// SIMATIC S7-200 project (STEP 7-Micro/WIN), CPU 226 CN REL 02.01

SYMBOL_TABLE 用户定义1
原点传感器检测          I0.0
右限位行程开关          I0.1
左限位行程开关          I0.2
机械手抬升下限检测        I0.3
机械手抬升上限检测        I0.4
机械手旋转左旋检测        I0.5
机械手旋转右旋检测        I0.6
机械手伸出检测          I0.7
机械手缩回检测          I1.0
机械手夹紧检测          I1.1
伺服报警             I1.2
按钮SB2            I2.4
按钮SB1            I2.5
急停               I2.6
全线速度             I2.7
初始状态检查           M0.0
回原点开始            M0.1
回原点完成            M0.2
正向点动             M0.3
反向点动             M0.4
双按键              M0.5
网络正常             M1.0
全线模式             M1.1
机械手复位            M1.2
准备就绪             M1.3
全线启动             M1.4
全线停止             M1.5
脉冲               Q0.0
方向               Q0.1
提升台上升电磁阀         Q0.3
回转气缸左旋电磁阀        Q0.4
回转气缸右旋电磁阀        Q0.5
手爪伸出电磁阀          Q0.6
手爪夹紧电磁阀          Q0.7
手爪放松电磁阀          Q1.0
黄色指示灯            Q1.5
绿色指示灯            Q1.6
红色指示灯            Q1.7
测试开始             S1.0
复位               V100.0
启动               V100.1
初始状态指示           V200.0
确认保存             V200.1
测试完成             V200.2
运行模式             V200.5
允许返回             V200.6
自动返回             V200.7
绿色警示灯            V1000.0
黄色警示灯            V1000.1
红色警示灯            V1000.2
各站红灯             V1000.3
供料请求             V1000.4
允许装配             V1000.5
允许加工             V1000.6
允许分拣             V1000.7
料不足_供料           V1020.2
缺料_供料            V1020.3
供料完成             V1020.4
料不足_装配           V1030.2
缺料_装配            V1030.3
装配完成             V1030.4
装配急停             V1030.5
故障无法修复           V1030.6
加工完成             V1040.2
停止完成             V1050.2
测试项              VB110
计划生产套件数          VB120
已生产套件数           VB1051
供料站位置            VD210
装配站位置            VD220
加工站位置            VD230
分拣站位置            VD240
当前绝对位置           VD250
当前速度             VD260
停止               V1001.0
END_SYMBOL_TABLE

ORGANIZATION_BLOCK 主程序:OB1
TITLE=程序注释
BEGIN
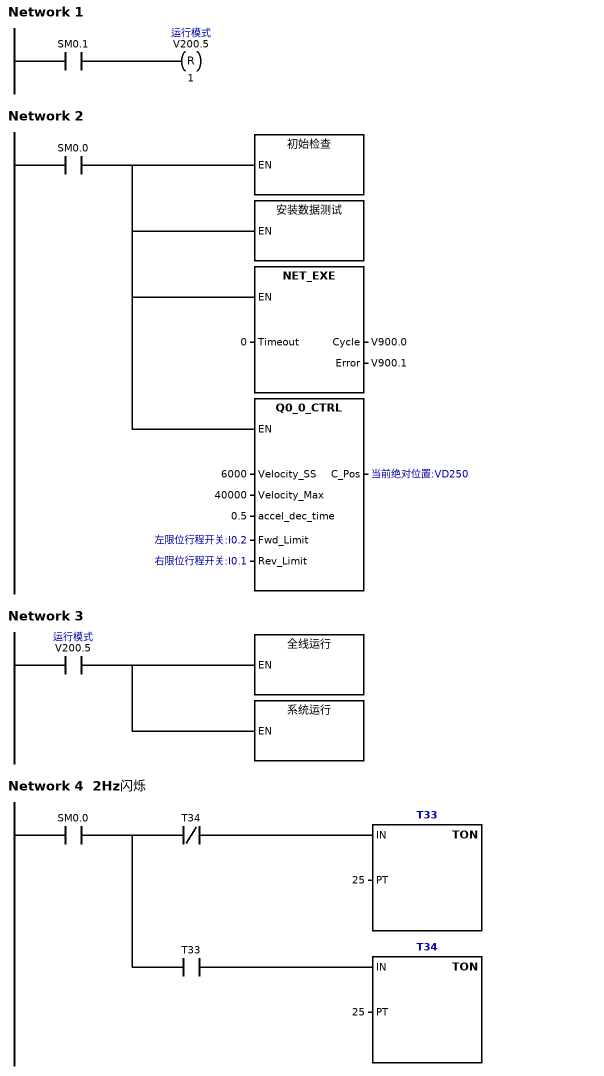
Network 1
LD     SM0.1
R      运行模式:V200.5, 1
Network 2
LD     SM0.0
CALL   初始检查:SBR0
CALL   安装数据测试:SBR8
CALL   NET_EXE:SBR11, 0, V900.0, V900.1
CALL   Q0_0_CTRL:SBR1, 6000, 40000, 0.5, 左限位行程开关:I0.2, 右限位行程开关:I0.1, 当前绝对位置:VD250
Network 3
LD     运行模式:V200.5
CALL   全线运行:SBR13
CALL   系统运行:SBR14
Network 4 // 2Hz闪烁
LD     SM0.0
LPS
AN     T34
TON    T33, 25
LPP
A      T33
TON    T34, 25
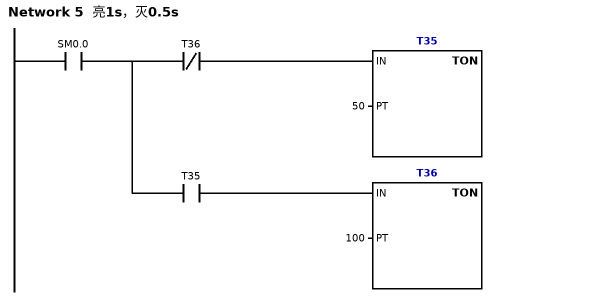
Network 5 // 亮1s，灭0.5s
LD     SM0.0
LPS
AN     T36
TON    T35, 50
LPP
A      T35
TON    T36, 100
END_ORGANIZATION_BLOCK

SUBROUTINE_BLOCK 初始检查:SBR0
TITLE=子程序注释
BEGIN
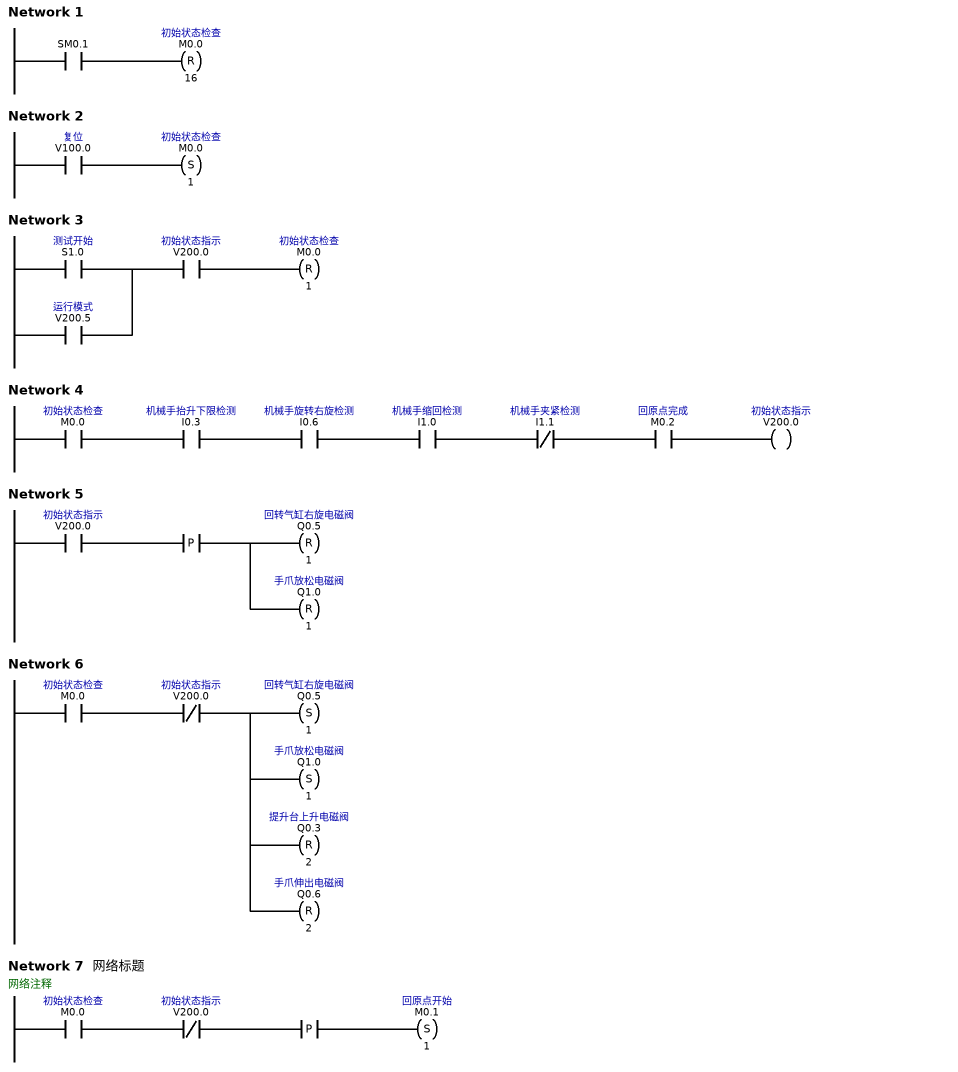
Network 1
LD     SM0.1
R      初始状态检查:M0.0, 16
Network 2
LD     复位:V100.0
S      初始状态检查:M0.0, 1
Network 3
LD     测试开始:S1.0
O      运行模式:V200.5
A      初始状态指示:V200.0
R      初始状态检查:M0.0, 1
Network 4
LD     初始状态检查:M0.0
A      机械手抬升下限检测:I0.3
A      机械手旋转右旋检测:I0.6
A      机械手缩回检测:I1.0
AN     机械手夹紧检测:I1.1
A      回原点完成:M0.2
=      初始状态指示:V200.0
Network 5
LD     初始状态指示:V200.0
EU
R      回转气缸右旋电磁阀:Q0.5, 1
R      手爪放松电磁阀:Q1.0, 1
Network 6
LD     初始状态检查:M0.0
AN     初始状态指示:V200.0
S      回转气缸右旋电磁阀:Q0.5, 1
S      手爪放松电磁阀:Q1.0, 1
R      提升台上升电磁阀:Q0.3, 2
R      手爪伸出电磁阀:Q0.6, 2
Network 7 // 网络标题
// 网络注释
LD     初始状态检查:M0.0
AN     初始状态指示:V200.0
EU
S      回原点开始:M0.1, 1
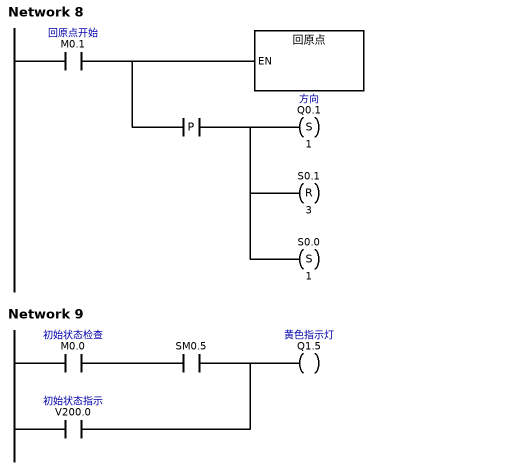
Network 8
LD     回原点开始:M0.1
CALL   回原点:SBR7
EU
S      方向:Q0.1, 1
R      S0.1, 3
S      S0.0, 1
Network 9
LD     初始状态检查:M0.0
A      SM0.5
O      初始状态指示:V200.0
=      黄色指示灯:Q1.5
END_SUBROUTINE_BLOCK

// SBR1: protected block, not included

// SBR2: protected block, not included

// SBR3: protected block, not included

// SBR4: protected block, not included

// SBR5: protected block, not included

// SBR6: protected block, not included

SUBROUTINE_BLOCK 回原点:SBR7
TITLE=子程序注释
BEGIN
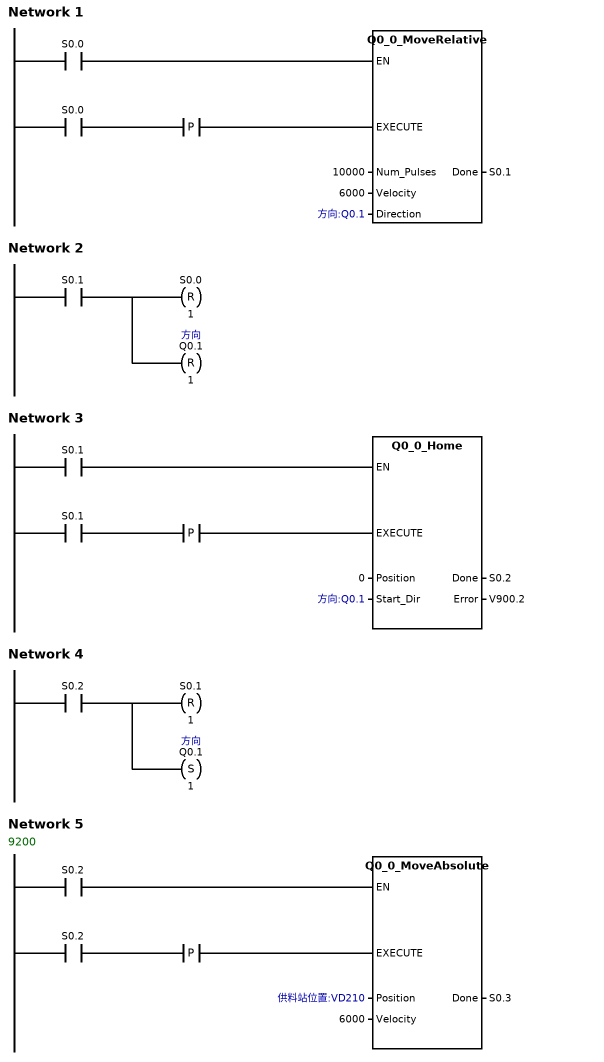
Network 1
LD     S0.0
=      L60.0
LD     S0.0
EU
=      L63.7
LD     L60.0
CALL   Q0_0_MoveRelative:SBR3, L63.7, 10000, 6000, 方向:Q0.1, S0.1
Network 2
LD     S0.1
R      S0.0, 1
R      方向:Q0.1, 1
Network 3
LD     S0.1
=      L60.0
LD     S0.1
EU
=      L63.7
LD     L60.0
CALL   Q0_0_Home:SBR5, L63.7, 0, 方向:Q0.1, S0.2, V900.2
Network 4
LD     S0.2
R      S0.1, 1
S      方向:Q0.1, 1
Network 5
// 9200
LD     S0.2
=      L60.0
LD     S0.2
EU
=      L63.7
LD     L60.0
CALL   Q0_0_MoveAbsolute:SBR4, L63.7, 供料站位置:VD210, 6000, S0.3
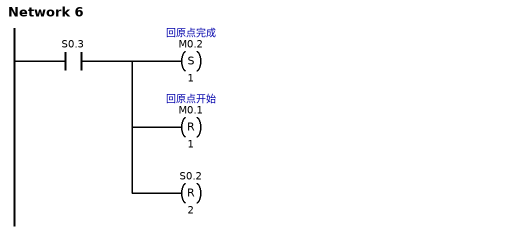
Network 6
LD     S0.3
S      回原点完成:M0.2, 1
R      回原点开始:M0.1, 1
R      S0.2, 2
Network 7 // 网络标题
// 网络注释
Network 9 // 网络标题
// 网络注释
END_SUBROUTINE_BLOCK

SUBROUTINE_BLOCK 安装数据测试:SBR8
TITLE=子程序注释
BEGIN
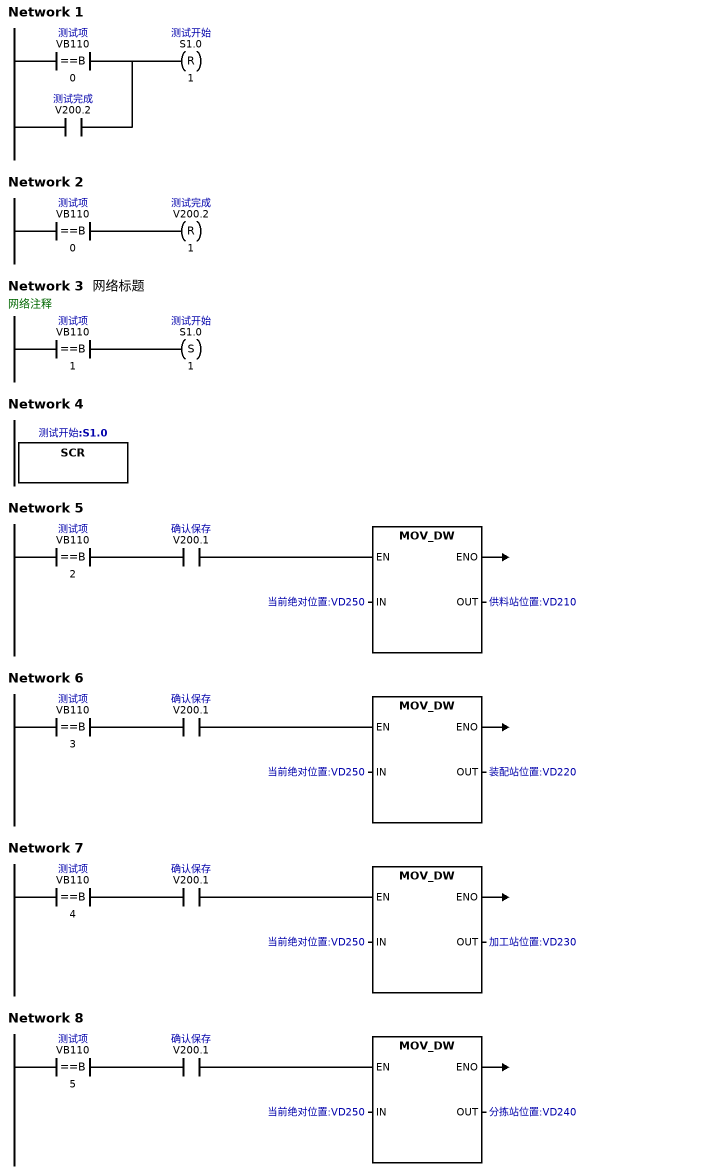
Network 1
LDB=   测试项:VB110, 0
O      测试完成:V200.2
R      测试开始:S1.0, 1
Network 2
LDB=   测试项:VB110, 0
R      测试完成:V200.2, 1
Network 3 // 网络标题
// 网络注释
LDB=   测试项:VB110, 1
S      测试开始:S1.0, 1
Network 4
LSCR   测试开始:S1.0
Network 5
LDB=   测试项:VB110, 2
A      确认保存:V200.1
MOVD   当前绝对位置:VD250, 供料站位置:VD210
Network 6
LDB=   测试项:VB110, 3
A      确认保存:V200.1
MOVD   当前绝对位置:VD250, 装配站位置:VD220
Network 7
LDB=   测试项:VB110, 4
A      确认保存:V200.1
MOVD   当前绝对位置:VD250, 加工站位置:VD230
Network 8
LDB=   测试项:VB110, 5
A      确认保存:V200.1
MOVD   当前绝对位置:VD250, 分拣站位置:VD240
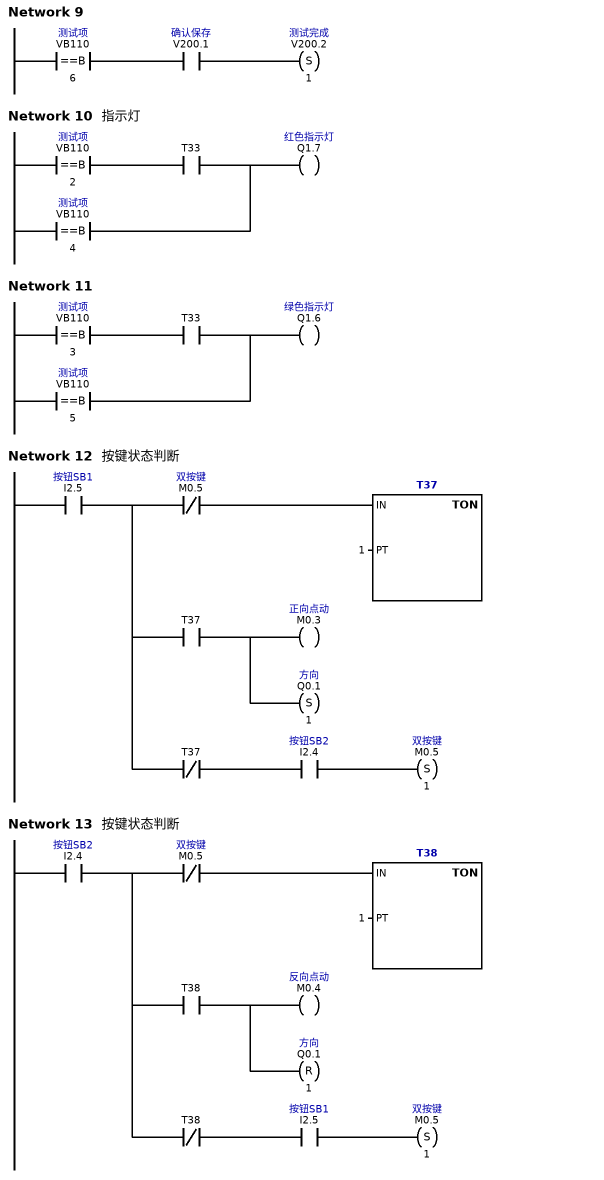
Network 9
LDB=   测试项:VB110, 6
A      确认保存:V200.1
S      测试完成:V200.2, 1
Network 10 // 指示灯
LDB=   测试项:VB110, 2
A      T33
OB=    测试项:VB110, 4
=      红色指示灯:Q1.7
Network 11
LDB=   测试项:VB110, 3
A      T33
OB=    测试项:VB110, 5
=      绿色指示灯:Q1.6
Network 12 // 按键状态判断
LD     按钮SB1:I2.5
LPS
AN     双按键:M0.5
TON    T37, 1
LRD
A      T37
=      正向点动:M0.3
S      方向:Q0.1, 1
LPP
AN     T37
A      按钮SB2:I2.4
S      双按键:M0.5, 1
Network 13 // 按键状态判断
LD     按钮SB2:I2.4
LPS
AN     双按键:M0.5
TON    T38, 1
LRD
A      T38
=      反向点动:M0.4
R      方向:Q0.1, 1
LPP
AN     T38
A      按钮SB1:I2.5
S      双按键:M0.5, 1
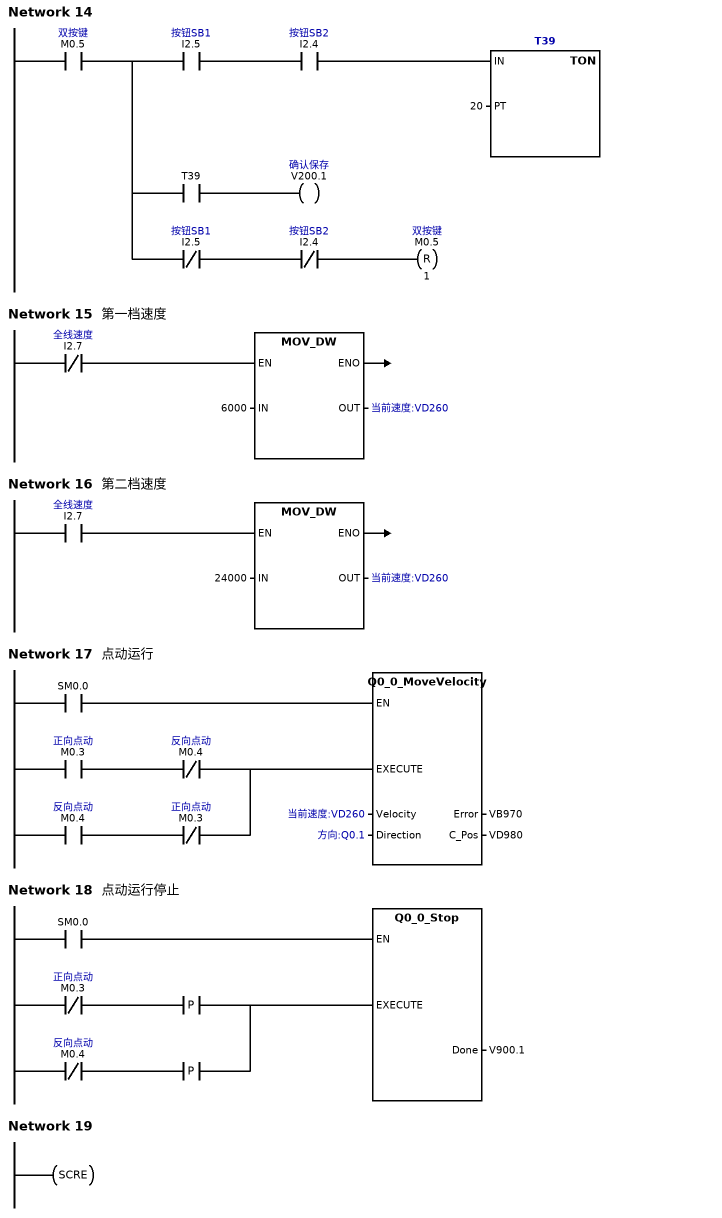
Network 14
LD     双按键:M0.5
LPS
A      按钮SB1:I2.5
A      按钮SB2:I2.4
TON    T39, 20
LRD
A      T39
=      确认保存:V200.1
LPP
AN     按钮SB1:I2.5
AN     按钮SB2:I2.4
R      双按键:M0.5, 1
Network 15 // 第一档速度
LDN    全线速度:I2.7
MOVD   6000, 当前速度:VD260
Network 16 // 第二档速度
LD     全线速度:I2.7
MOVD   24000, 当前速度:VD260
Network 17 // 点动运行
LD     SM0.0
=      L60.0
LD     正向点动:M0.3
AN     反向点动:M0.4
LD     反向点动:M0.4
AN     正向点动:M0.3
OLD
=      L63.7
LD     L60.0
CALL   Q0_0_MoveVelocity:SBR9, L63.7, 当前速度:VD260, 方向:Q0.1, VB970, VD980
Network 18 // 点动运行停止
LD     SM0.0
=      L60.0
LDN    正向点动:M0.3
EU
LDN    反向点动:M0.4
EU
OLD
=      L63.7
LD     L60.0
CALL   Q0_0_Stop:SBR10, L63.7, V900.1
Network 19
SCRE
END_SUBROUTINE_BLOCK

// SBR9: protected block, not included

// SBR10: protected block, not included

// SBR11: protected block, not included

SUBROUTINE_BLOCK 全线运行:SBR13
TITLE=
BEGIN
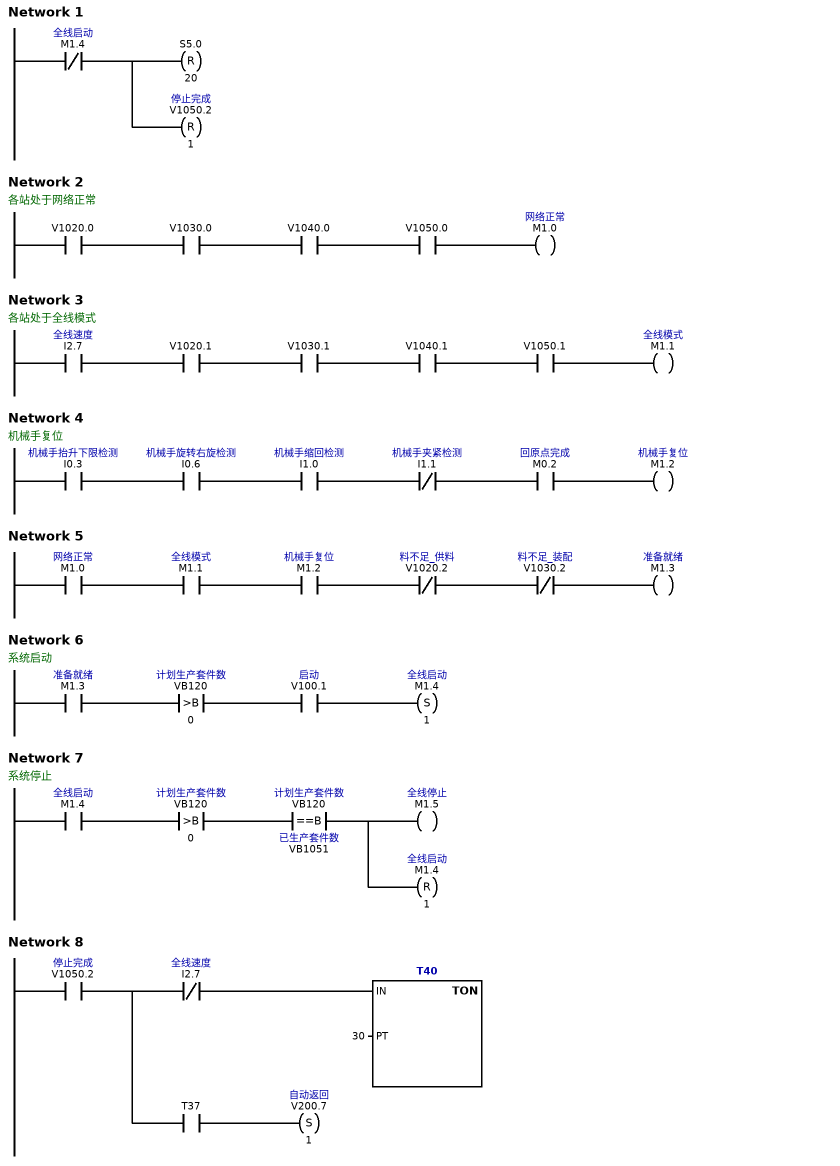
Network 1
LDN    全线启动:M1.4
R      S5.0, 20
R      停止完成:V1050.2, 1
Network 2
// 各站处于网络正常
LD     V1020.0
A      V1030.0
A      V1040.0
A      V1050.0
=      网络正常:M1.0
Network 3
// 各站处于全线模式
LD     全线速度:I2.7
A      V1020.1
A      V1030.1
A      V1040.1
A      V1050.1
=      全线模式:M1.1
Network 4
// 机械手复位
LD     机械手抬升下限检测:I0.3
A      机械手旋转右旋检测:I0.6
A      机械手缩回检测:I1.0
AN     机械手夹紧检测:I1.1
A      回原点完成:M0.2
=      机械手复位:M1.2
Network 5
LD     网络正常:M1.0
A      全线模式:M1.1
A      机械手复位:M1.2
AN     料不足_供料:V1020.2
AN     料不足_装配:V1030.2
=      准备就绪:M1.3
Network 6
// 系统启动
LD     准备就绪:M1.3
AB>    计划生产套件数:VB120, 0
A      启动:V100.1
S      全线启动:M1.4, 1
Network 7
// 系统停止
LD     全线启动:M1.4
AB>    计划生产套件数:VB120, 0
AB=    计划生产套件数:VB120, 已生产套件数:VB1051
=      全线停止:M1.5
R      全线启动:M1.4, 1
Network 8
LD     停止完成:V1050.2
LPS
AN     全线速度:I2.7
TON    T40, 30
LPP
A      T37
S      自动返回:V200.7, 1
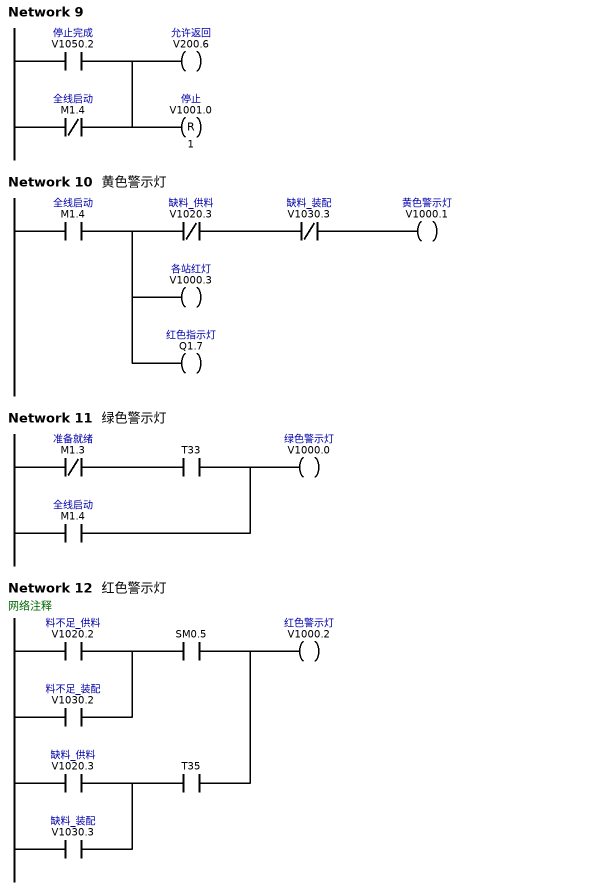
Network 9
LD     停止完成:V1050.2
ON     全线启动:M1.4
=      允许返回:V200.6
R      停止:V1001.0, 1
Network 10 // 黄色警示灯
LD     全线启动:M1.4
LPS
AN     缺料_供料:V1020.3
AN     缺料_装配:V1030.3
=      黄色警示灯:V1000.1
LRD
=      各站红灯:V1000.3
LPP
=      红色指示灯:Q1.7
Network 11 // 绿色警示灯
LDN    准备就绪:M1.3
A      T33
O      全线启动:M1.4
=      绿色警示灯:V1000.0
Network 12 // 红色警示灯
// 网络注释
LD     料不足_供料:V1020.2
O      料不足_装配:V1030.2
A      SM0.5
LD     缺料_供料:V1020.3
O      缺料_装配:V1030.3
A      T35
OLD
=      红色警示灯:V1000.2
END_SUBROUTINE_BLOCK

SUBROUTINE_BLOCK 系统运行:SBR14
TITLE=子程序注释
BEGIN
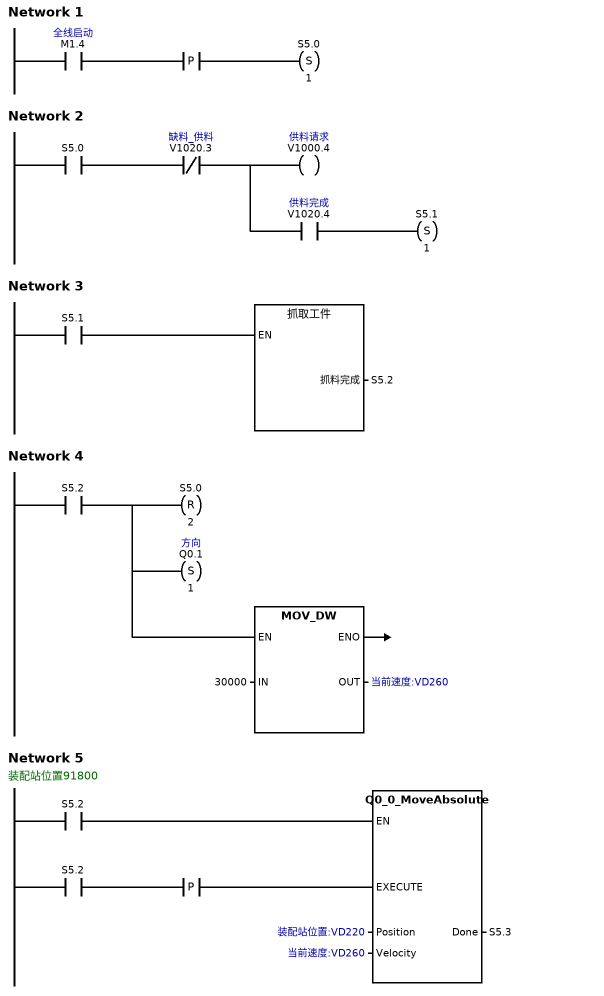
Network 1
LD     全线启动:M1.4
EU
S      S5.0, 1
Network 2
LD     S5.0
AN     缺料_供料:V1020.3
=      供料请求:V1000.4
A      供料完成:V1020.4
S      S5.1, 1
Network 3
LD     S5.1
CALL   抓取工件:SBR15, S5.2
Network 4
LD     S5.2
R      S5.0, 2
S      方向:Q0.1, 1
MOVD   30000, 当前速度:VD260
Network 5
// 装配站位置91800
LD     S5.2
=      L60.0
LD     S5.2
EU
=      L63.7
LD     L60.0
CALL   Q0_0_MoveAbsolute:SBR4, L63.7, 装配站位置:VD220, 当前速度:VD260, S5.3
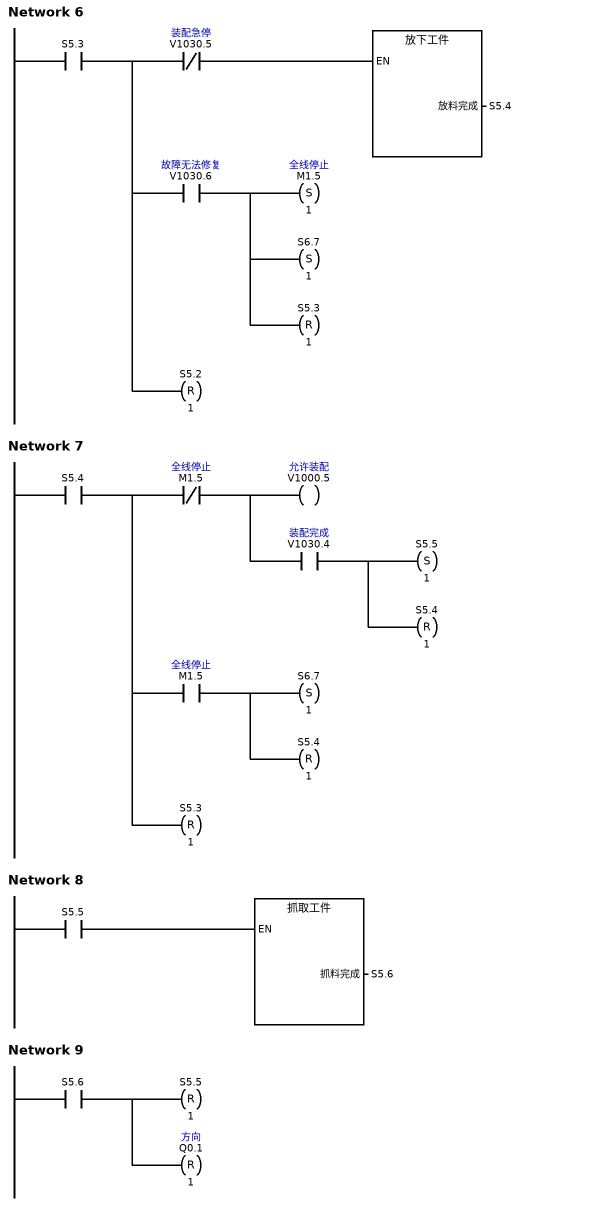
Network 6
LD     S5.3
LPS
AN     装配急停:V1030.5
CALL   放下工件:SBR16, S5.4
LRD
A      故障无法修复:V1030.6
S      全线停止:M1.5, 1
S      S6.7, 1
R      S5.3, 1
LPP
R      S5.2, 1
Network 7
LD     S5.4
LPS
AN     全线停止:M1.5
=      允许装配:V1000.5
A      装配完成:V1030.4
S      S5.5, 1
R      S5.4, 1
LPP
LPS
A      全线停止:M1.5
S      S6.7, 1
R      S5.4, 1
LPP
R      S5.3, 1
Network 8
LD     S5.5
CALL   抓取工件:SBR15, S5.6
Network 9
LD     S5.6
R      S5.5, 1
R      方向:Q0.1, 1
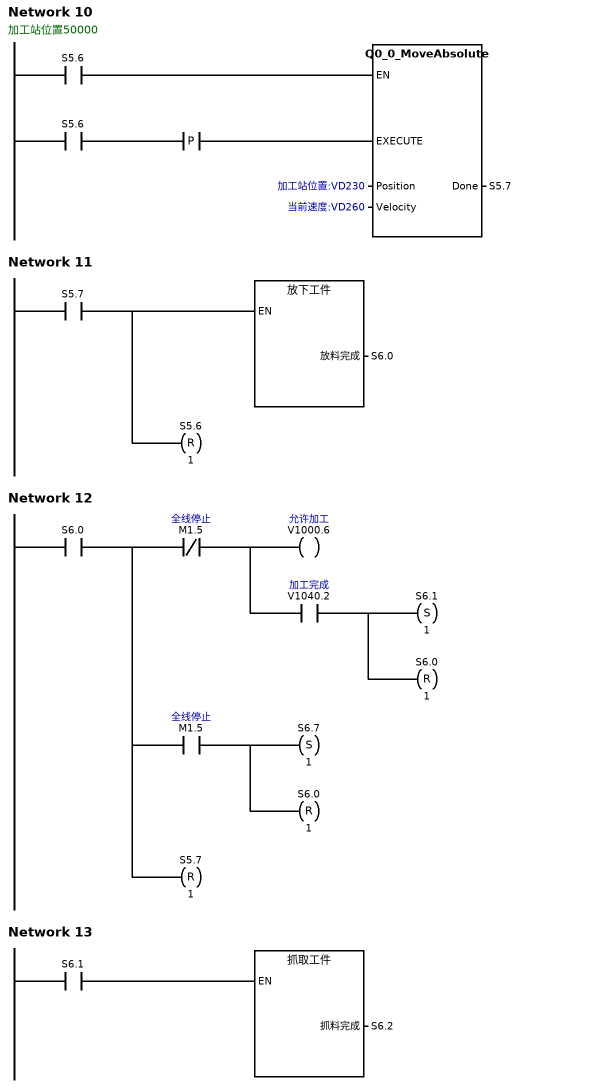
Network 10
// 加工站位置50000
LD     S5.6
=      L60.0
LD     S5.6
EU
=      L63.7
LD     L60.0
CALL   Q0_0_MoveAbsolute:SBR4, L63.7, 加工站位置:VD230, 当前速度:VD260, S5.7
Network 11
LD     S5.7
CALL   放下工件:SBR16, S6.0
R      S5.6, 1
Network 12
LD     S6.0
LPS
AN     全线停止:M1.5
=      允许加工:V1000.6
A      加工完成:V1040.2
S      S6.1, 1
R      S6.0, 1
LPP
LPS
A      全线停止:M1.5
S      S6.7, 1
R      S6.0, 1
LPP
R      S5.7, 1
Network 13
LD     S6.1
CALL   抓取工件:SBR15, S6.2
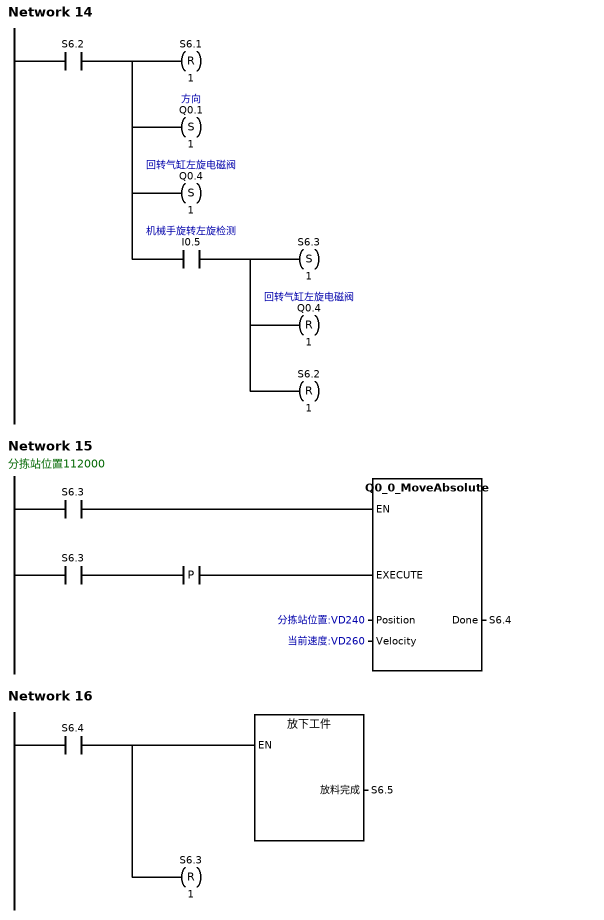
Network 14
LD     S6.2
R      S6.1, 1
S      方向:Q0.1, 1
S      回转气缸左旋电磁阀:Q0.4, 1
A      机械手旋转左旋检测:I0.5
S      S6.3, 1
R      回转气缸左旋电磁阀:Q0.4, 1
R      S6.2, 1
Network 15
// 分拣站位置112000
LD     S6.3
=      L60.0
LD     S6.3
EU
=      L63.7
LD     L60.0
CALL   Q0_0_MoveAbsolute:SBR4, L63.7, 分拣站位置:VD240, 当前速度:VD260, S6.4
Network 16
LD     S6.4
CALL   放下工件:SBR16, S6.5
R      S6.3, 1
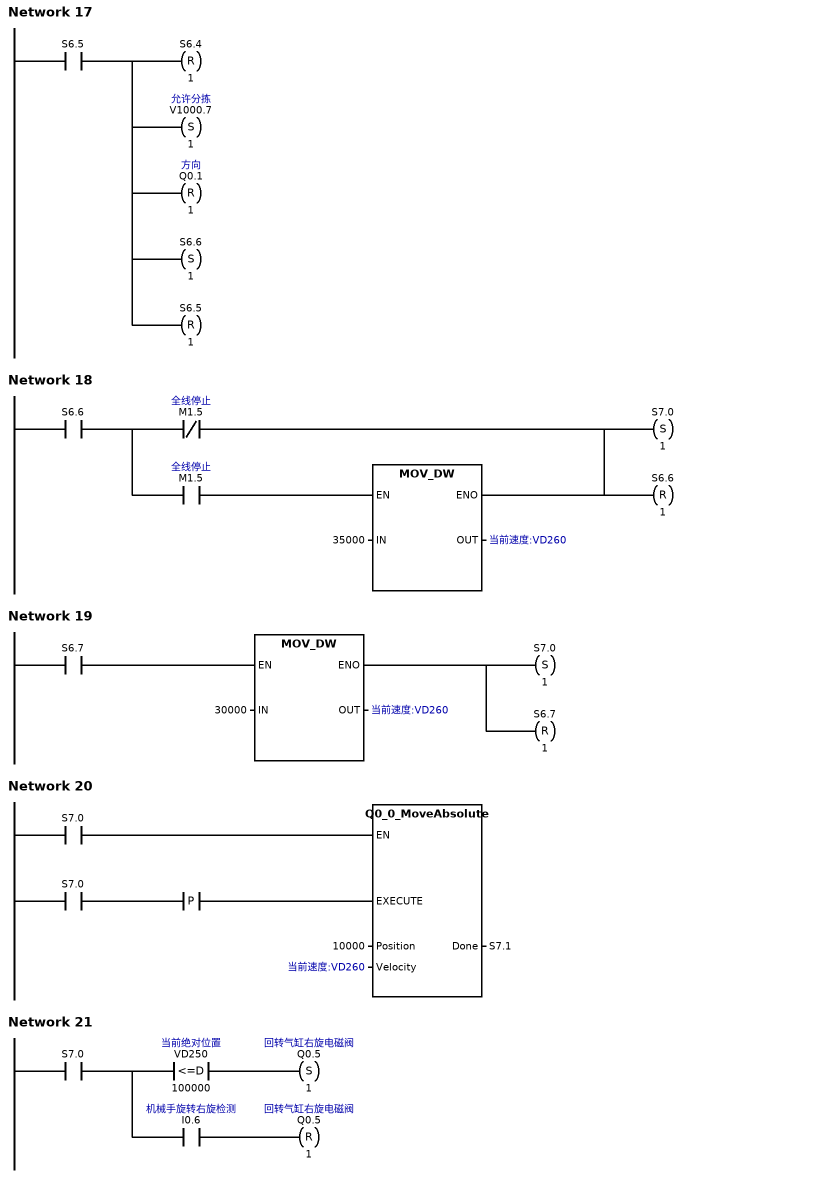
Network 17
LD     S6.5
R      S6.4, 1
S      允许分拣:V1000.7, 1
R      方向:Q0.1, 1
S      S6.6, 1
R      S6.5, 1
Network 18
LD     S6.6
LPS
AN     全线停止:M1.5
=      L63.7
LPP
A      全线停止:M1.5
MOVD   35000, 当前速度:VD260
AENO
O      L63.7
S      S7.0, 1
R      S6.6, 1
Network 19
LD     S6.7
MOVD   30000, 当前速度:VD260
AENO
S      S7.0, 1
R      S6.7, 1
Network 20
LD     S7.0
=      L60.0
LD     S7.0
EU
=      L63.7
LD     L60.0
CALL   Q0_0_MoveAbsolute:SBR4, L63.7, 10000, 当前速度:VD260, S7.1
Network 21
LD     S7.0
LPS
AD<=   当前绝对位置:VD250, 100000
S      回转气缸右旋电磁阀:Q0.5, 1
LPP
A      机械手旋转右旋检测:I0.6
R      回转气缸右旋电磁阀:Q0.5, 1
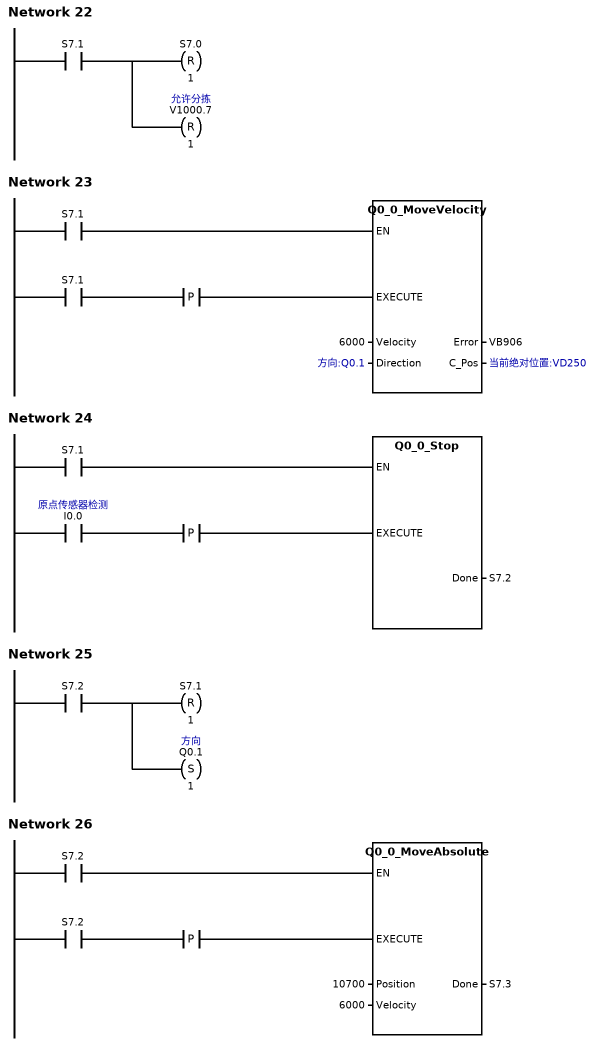
Network 22
LD     S7.1
R      S7.0, 1
R      允许分拣:V1000.7, 1
Network 23
LD     S7.1
=      L60.0
LD     S7.1
EU
=      L63.7
LD     L60.0
CALL   Q0_0_MoveVelocity:SBR9, L63.7, 6000, 方向:Q0.1, VB906, 当前绝对位置:VD250
Network 24
LD     S7.1
=      L60.0
LD     原点传感器检测:I0.0
EU
=      L63.7
LD     L60.0
CALL   Q0_0_Stop:SBR10, L63.7, S7.2
Network 25
LD     S7.2
R      S7.1, 1
S      方向:Q0.1, 1
Network 26
LD     S7.2
=      L60.0
LD     S7.2
EU
=      L63.7
LD     L60.0
CALL   Q0_0_MoveAbsolute:SBR4, L63.7, 10700, 6000, S7.3
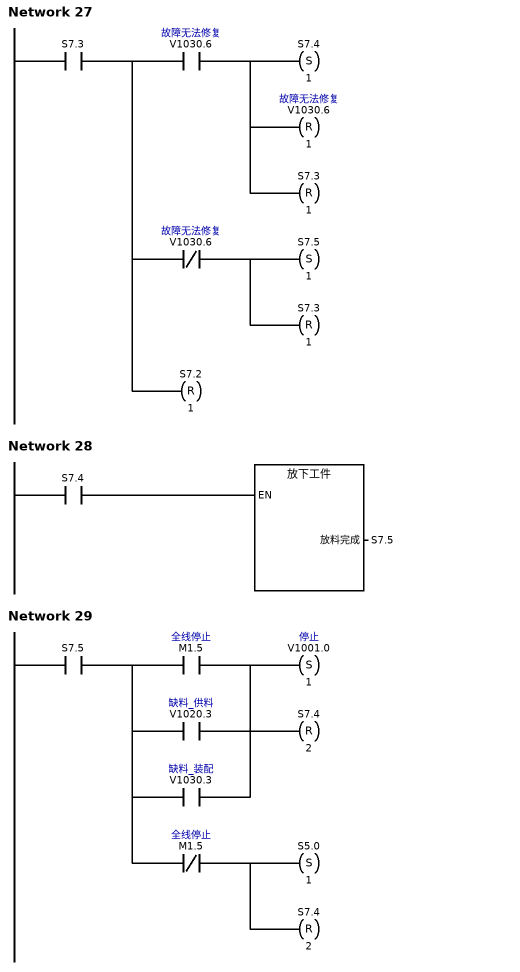
Network 27
LD     S7.3
LPS
A      故障无法修复:V1030.6
S      S7.4, 1
R      故障无法修复:V1030.6, 1
R      S7.3, 1
LRD
AN     故障无法修复:V1030.6
S      S7.5, 1
R      S7.3, 1
LPP
R      S7.2, 1
Network 28
LD     S7.4
CALL   放下工件:SBR16, S7.5
Network 29
LD     S7.5
LPS
LD     全线停止:M1.5
O      缺料_供料:V1020.3
O      缺料_装配:V1030.3
ALD
S      停止:V1001.0, 1
R      S7.4, 2
LPP
AN     全线停止:M1.5
S      S5.0, 1
R      S7.4, 2
END_SUBROUTINE_BLOCK

SUBROUTINE_BLOCK 抓取工件:SBR15
TITLE=子程序注释
VAR_OUTPUT
抓料完成:BOOL;	// L0.0 
END_VAR
BEGIN
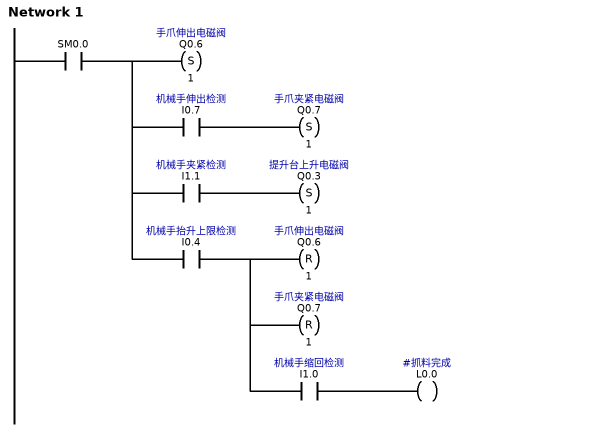
Network 1
LD     SM0.0
LPS
S      手爪伸出电磁阀:Q0.6, 1
A      机械手伸出检测:I0.7
S      手爪夹紧电磁阀:Q0.7, 1
LRD
A      机械手夹紧检测:I1.1
S      提升台上升电磁阀:Q0.3, 1
LPP
A      机械手抬升上限检测:I0.4
R      手爪伸出电磁阀:Q0.6, 1
R      手爪夹紧电磁阀:Q0.7, 1
A      机械手缩回检测:I1.0
=      #抓料完成:L0.0
Network 2 // 网络标题
// 网络注释
END_SUBROUTINE_BLOCK
